(* IEC 61131-3 sources: kns-port-domestic/targets/astra/src/POUs/Generated/PRG_ApplyProjectCfg, 1 file *)

(* ---- PRG_ApplyProjectCfg.decl.st ---- *)
// AUTO-GENERATED by iolistgen 0.2.0 — не редактировать; источник: 03_io_list.csv
// SHA-256 перечня 06336d13c4b2; генератор st-codesys
// Назначение: «применить уставки проекта»: копирует GVL_CfgProject.st<DEV>Cfg в GVL_Persist.st<DEV>Cfg; Retain
// устройств не меняется (контракт plc-process-lib 18.3, правило 2). Вызывается из PRG_Devices по команде
// GVL_Hmi.xApplyProjectCfg или из логики станции
// Автор:      iolistgen (генератор по перечню сигналов); перечень 03_io_list.csv
// Версия:     iolistgen 0.2.0
// Документ:   docs/03_io_list.md
PROGRAM PRG_ApplyProjectCfg
VAR
END_VAR
